// TIA Portal V18 export
VAR_GLOBAL   // PLC tag table "Default tag table"
   System_Byte AT %MB1 : Byte;
   FirstScan AT %M1.0 : Bool;
   DiagStatusUpdate AT %M1.1 : Bool;
   AlwaysTRUE AT %M1.2 : Bool;
   AlwaysFALSE AT %M1.3 : Bool;
   Clock_Byte AT %MB0 : Byte;
   Clock_10Hz AT %M0.0 : Bool;
   Clock_5Hz AT %M0.1 : Bool;
   "Clock_2.5Hz" AT %M0.2 : Bool;
   Clock_2Hz AT %M0.3 : Bool;
   "Clock_1.25Hz" AT %M0.4 : Bool;
   Clock_1Hz AT %M0.5 : Bool;
   "Clock_0.625Hz" AT %M0.6 : Bool;
   "Clock_0.5Hz" AT %M0.7 : Bool;
   Tag_MotorOnOff AT %Q0.0 : Bool;
   analogInput_1 AT %IW64 : Int;
   analogInput_2 AT %IW66 : Int;
END_VAR
VAR_GLOBAL CONSTANT   // user constants
   ReadMonitorParams : Int := 0;
   ReadCommandRegs : Int := 1;
   WriteMotorOnOff : Int := 3;
   WriteFrequencySetpoint : Int := 4;
   WriteSpeedSourceSelect : Int := 5;
   ReadAlarmHistory : Int := 6;
   ReadAlarm : Int := 2;
   alarm_UV1 : Int := 0;
   alarm_UV3 : Int := 1;
   alarm_SC : Int := 2;
   alarm_OC : Int := 3;
   alarm_OV : Int := 4;
   alarm_OH : Int := 5;
   alarm_OL1 : Int := 6;
   alarm_OL2 : Int := 7;
   alarm_CPF03 : Int := 8;
   alarm_StopMod_LowZPT : Int := 9;
   alarm_StopMod_HighZPT : Int := 10;
   alarm_StopMod_OverheatingRadiator : Int := 11;
   alarm_StopMod_bb : Int := 12;
   alarm_CTER : Int := 13;
   alarm_FBL : Int := 14;
   alarm_ES : Int := 15;
   alarm_STP0 : Int := 16;
   alarm_STP1 : Int := 17;
   alarm_STP2 : Int := 18;
   WriteResetAlarm : Int := 7;
END_VAR
